(* IEC 61131-3 sources: 89152_FlorisHendrix_AfstudeerProject/89152_FlorisHendrix_ExamenProject/Stations/Terminal/HMI/Network/NewAgeSettings, 1 file *)

(* ---- ONE_NewAgeSettings_Table.st ---- *)
#define OBJECTS_CONFIG

//Define part of class USB_DataExchange
#define USB_DATA_CMD                  16#10
#define USB_DataExchangeBase_Timeout  10ms
#define continue goto LABEL_continue
#include "..\..\Source\interfaces\lsl_st_Usb.h"
//Define part of class DisplaySettings
#define DISPLAYSETTINGS_OS_STARTVERSION_SALAMANDER 0x9100  // salamder starts with v 9.1.00

#define DISPLAYSETTINGS_GRAPHIX_MAX_BRIGHTNESS  255 //(2^8-1) = 255
#define DISPLAYSETTINGS_USB_MAX_BRIGHTNESS      255 //(2^8-1) = 255
#define DISPLAYSETTINGS_MIN_BRIGHTNESS_INPUT      0
#define DISPLAYSETTINGS_MAX_BRIGHTNESS_INPUT    100

#define DISPLAYSETTINGS_MIN_PWM_INPUT          0
#define DISPLAYSETTINGS_MAX_PWM_INPUT          100
#define DISPLAYSETTINGS_PWM_PERIODE_TIME       10000

#define DISPLAYSETTINGS_USB_REQ_TIMER_UP 1000

#define DISPLAYSETTINGS_USB_INIT_ERROR    -1

#define DISPLAYSETTINGS_BRIGHTNESS_ERROR    -1

#define DISPLAYSETTINGS_TASKOBJECT_NOT_FOUND    -5

#define DISPLAYSETTINGS_STATE_OK                0

#define DISPLAYSETTINGS_BACKGROUNDTASK_ERROR    -1
#define DISPLAYSETTINGS_CAN_OBJECT_ERROR        -2
#define DISPLAYSETTINGS_GRAPHIX_ERROR           -3
#define DISPLAYSETTINGS_PSOC_ERROR               -4

#define DISPLAYSETTINGS_BACKLIGHT_SWITCHOFF_TIME 1000 //1 second
#include "..\..\Source\interfaces\lsl_st_kernel.h"
#include "..\..\Source\interfaces\lsl_st_pci.h"
#include "..\..\Source\interfaces\lsl_st_pwm.h"
#include "..\..\Source\interfaces\lsl_st_gpio.h"
#include "..\..\Source\interfaces\lsl_st_screensaver.h"
//Define part of class KeyPadANumStdTemplate
#define KEY_LAYOUT_LINE_1   2#11111111110
#define KEY_LAYOUT_LINE_2   2#11111111110
#define KEY_LAYOUT_LINE_3   2#01111111110
#define KEY_LAYOUT_LINE_4   2#00000000111

#define KEYPAD_ANUM_BUTTON_WIDTH      60
#define KEYPAD_ANUM_BUTTON_HEIGHT     60

#define KEYPAD_ANUM_BUTTON_XOFF       5
#define KEYPAD_ANUM_BUTTON_YOFF       85

#define KEYPAD_ANUM_WIDTH             680
#define KEYPAD_ANUM_HEIGHT            350

#define KEYPAD_ANUM_INPUT_XOFF        5
#define KEYPAD_ANUM_INPUT_YOFF        45
#define KEYPAD_ANUM_INPUT_HEIGHT      30

#define KEYPAD_ANUM_TITLE_XOFF        5
#define KEYPAD_ANUM_TITLE_YOFF        5
#define KEYPAD_ANUM_TITLE_HEIGHT      30

#define KEYPAD_ANUM_ESC_WIDTH         30
//Define part of class KeyPadNumStdTemplate
#define KEYPAD_NUM_BUTTON_WIDTH       80
#define KEYPAD_NUM_BUTTON_HEIGHT      80

#define KEYPAD_NUM_BUTTON_XOFF        5
#define KEYPAD_NUM_BUTTON_YOFF        105

#define KEYPAD_NUM_WIDTH              330
#define KEYPAD_NUM_HEIGHT             435

#define KEYPAD_NUM_INPUT_XOFF         5
#define KEYPAD_NUM_INPUT_YOFF         45
#define KEYPAD_NUM_INPUT_HEIGHT       30

#define KEYPAD_NUM_TITLE_XOFF         7
#define KEYPAD_NUM_TITLE_YOFF         5
#define KEYPAD_NUM_TITLE_HEIGHT       30

#define KEYPAD_NUM_LIMIT_XOFF         5
#define KEYPAD_NUM_LIMIT_YOFF         80
#define KEYPAD_NUM_LIMIT_WIDTH        80
#define KEYPAD_NUM_LIMIT_HEIGTH       20

#define KEYPAD_NUM_UNIT_WIDTH         70
#define KEYPAD_NUM_UNIT_HEIGTH        20

#define KEYPAD_NUM_ESC_WIDTH          30
//Define part of class SystemLogging
//texts for indicating type of loginformation
#define LOG_TYPE_ERROR    ("ERROR:")
#define LOG_TYPE_WARNING  ("WARNING:")
#define LOG_TYPE_DEBUG    ("DEBUG:")
#define LOG_TYPE_INFO     ("INFO:")
//Define part of class TouchCalib
// Default-Settings for the Touch-Calibration
//-------------------------------------------------------------------------------------------------

#define   TouchCalib_UDCVersion                                         1
#define   TouchCalib_NoAnything                                         2

#define   TouchCalib_TextTouchScreen                                    "Please touch the screen to start!"
#define   TouchCalib_TextTouchCrosshair                                 "Please touch the crosshair!"
#define   TouchCalib_TextCalibSuccessful                                "Calibration successful! Please touch the screen to continue."
#define   TouchCalib_TextCalibFailed                                    "Calibration failed! Please touch the screen to calibrate again."
#define   TouchCalib_TextNextScreen                                     "Calibration successful! Please touch the NEXT device to continue."

#define   TouchCalib_TextIdxTouchScreen                                 0
#define   TouchCalib_TextIdxTouchCrosshair                              1
#define   TouchCalib_TextIdxCalibSuccessful                             2
#define   TouchCalib_TextIdxCalibFailed                                 3
#define   TouchCalib_TextIdxNextScreen                                  4

#define   TouchCalib_StdTextAttrib                                      T_SOLID OR T_COPY OR T_PROP

#define   TouchCalib_CrosshairSize                                      40                                            // The length and width of the crosshair (if no image is chosen) [pixel]

#define   TouchCalib_MinTimeBewtweenTouchEvent                         100 ms

FUNCTION GLOBAL TAB ONE_NewAgeSettings
-1$UINT, 0$UINT,
1$UINT, 0$UINT,

15$UDINT,
TO_UDINT(3788417926), "_Global", 0$UINT, 15$UINT, 0$UINT,
TO_UDINT(1108585033), "_LanguageSelection", 0$UINT, 5$UINT, 1$UINT,
TO_UDINT(2980745877), "_MyIO", 0$UINT, 3$UINT, 0$UINT,
TO_UDINT(3599188277), "_Screen", 0$UINT, 3$UINT, 0$UINT,
TO_UDINT(3043040051), "_ScrollArea", 0$UINT, 15$UINT, 0$UINT,
TO_UDINT(2779823616), "_ScrollArea2", 0$UINT, 8$UINT, 0$UINT,
TO_UDINT(3306153856), "DisplaySettings", 1$UINT, 39$UINT, 1$UINT,
TO_UDINT(1679073929), "KeyPadANumStdTemplate", 3$UINT, 0$UINT, 1$UINT,
TO_UDINT(980817768), "KeyPadImagesStdTemplate", 2$UINT, 0$UINT, 2$UINT,
TO_UDINT(1267823535), "KeyPadNumStdTemplate", 1$UINT, 0$UINT, 1$UINT,
TO_UDINT(1903583397), "Ram", 1$UINT, 3$UINT, 1$UINT,
TO_UDINT(3719262472), "ScreenSaver", 1$UINT, 13$UINT, 1$UINT,
TO_UDINT(90452573), "SystemLogging", 1$UINT, 5$UINT, 1$UINT,
TO_UDINT(627189056), "TouchCalib", 1$UINT, 4$UINT, 1$UINT,
TO_UDINT(1659734526), "USB_DataExchange", 1$UINT, 14$UINT, 0$UINT,

_NO_ATTR, TO_UDINT(2359166249), "_LANGUAGESELECTION1",

1$UINT, TO_UDINT(474634808), "SCREENSAVER1\DISPLAYSETTINGS",

_NO_ATTR, TO_UDINT(1679073929), "KEYPADANUMSTDTEMPLATE",

1$UINT, TO_UDINT(860932433), "KEYPADANUMSTDTEMPLATE\KEYPADIMG",
1$UINT, TO_UDINT(1346448759), "KEYPADNUMSTDTEMPLATE\KEYPADIMG",

_NO_ATTR, TO_UDINT(1267823535), "KEYPADNUMSTDTEMPLATE",

_NO_ATTR, TO_UDINT(2623333383), "CLEANSCREENTIME",

_NO_ATTR, TO_UDINT(2379925748), "SCREENSAVER1",

_NO_ATTR, TO_UDINT(2516821708), "SYSTEMLOGGING1",

_NO_ATTR, TO_UDINT(4112894978), "TOUCHCALIB1",

//Internal connections
0$UDINT,
3$UDINT,
TO_UDINT(2), "KeyPadImg", TO_UDINT(3),
TO_UDINT(5), "KeyPadImg", TO_UDINT(4),
TO_UDINT(7), "DisplaySettings", TO_UDINT(1),
0$UDINT,
0$UDINT,

//Initialization values
0$UDINT,
18$UDINT,
TO_UDINT(0), "LineWidth", TO_UDINT(70),//|NewAgeSettings._LanguageSelection1.LineWidth;
TO_UDINT(0), "LineHighness", TO_UDINT(30),//|NewAgeSettings._LanguageSelection1.LineHighness;
TO_UDINT(0), "ExtendedScrollBar", TO_UDINT(0),//|NewAgeSettings._LanguageSelection1.ExtendedScrollBar;
TO_UDINT(0), "Config", TO_UDINT(3),//|NewAgeSettings._LanguageSelection1.Config;
TO_UDINT(1), "Brightness", TO_UDINT(100),//|NewAgeSettings.ScreenSaver1\DisplaySettings.Brightness;
TO_UDINT(1), "ScreensaverTime", TO_UDINT(60),//|NewAgeSettings.ScreenSaver1\DisplaySettings.ScreensaverTime;
TO_UDINT(2), "No", TO_UDINT(_WIN_EDITOR_ANUMERIC),//|NewAgeSettings.KeyPadANumStdTemplate.No;
TO_UDINT(2), "ImA", TO_UDINT(ImA_Window),//|NewAgeSettings.KeyPadANumStdTemplate.ImA;
TO_UDINT(5), "No", TO_UDINT(_WIN_EDITOR_NUMERIC),//|NewAgeSettings.KeyPadNumStdTemplate.No;
TO_UDINT(5), "ImA", TO_UDINT(IMA_WINDOW),//|NewAgeSettings.KeyPadNumStdTemplate.ImA;
TO_UDINT(6), "", TO_UDINT(5),//|NewAgeSettings.CleanScreenTime.Data;
TO_UDINT(7), "sDelayScreenSaver", TO_UDINT(0),//|NewAgeSettings.ScreenSaver1.sDelayScreenSaver;
TO_UDINT(7), "sDelayBacklight", TO_UDINT(0),//|NewAgeSettings.ScreenSaver1.sDelayBacklight;
TO_UDINT(7), "BrightnessMinStart", TO_UDINT(20),//|NewAgeSettings.ScreenSaver1.BrightnessMinStart;
TO_UDINT(8), "ExtLoggingActive", TO_UDINT(TRUE),//|NewAgeSettings.SystemLogging1.ExtLoggingActive;
TO_UDINT(8), "ActivateTrace", TO_UDINT(0),//|NewAgeSettings.SystemLogging1.ActivateTrace;
TO_UDINT(9), "SelectOrderNo", TO_UDINT(-1),//|NewAgeSettings.TouchCalib1.SelectOrderNo;
TO_UDINT(9), "Tolerance", TO_UDINT(20),//|NewAgeSettings.TouchCalib1.Tolerance;

//Symbolic initialization values
0$UDINT,
0$UDINT,

//Initialization of string values
0$UDINT,
0$UDINT,

//Configuration of tasks (RealTime, Cyclic, Background)
0$UDINT,
0$UDINT,

0$UDINT,
0$UDINT,

0$UDINT,
1$UDINT,
TO_UDINT(1), (-1)$UDINT, 4194303$DINT, 	//SCREENSAVER1\DISPLAYSETTINGS

//External connections
0$UDINT,
5$UDINT,
TO_UDINT(0), "Lse", C_DIR, TO_UDINT(299963966), "Lse","Lse",
TO_UDINT(2), "Lse", C_DIR, TO_UDINT(299963966), "Lse","Lse",
TO_UDINT(5), "Lse", C_DIR, TO_UDINT(299963966), "Lse","Lse",
TO_UDINT(7), "Lse", C_DIR, TO_UDINT(299963966), "Lse","Lse",
TO_UDINT(9), "Lse", C_DIR, TO_UDINT(299963966), "Lse","Lse",

//Magic internal connections
0$UDINT,
0$UDINT,

//Configuration of timeslots of tasks (RealTime, Cyclic)
#ifdef __LSLLDR_TIMESLOTS__
0$UDINT,
0$UDINT,

0$UDINT,
0$UDINT,

#endif //__LSLLDR_TIMESLOTS__

//MultiMaster connections
#ifdef __LSLLDR_MULTIMASTER__
0$UDINT,
0$UDINT,
#endif //__LSLLDR_MULTIMASTER__

//Configuration for task ID (RealTime, CyclicTime)
#ifdef __LSLLDR_TASKID__
"\\\\TASKS2  "
0$UDINT,
0$UDINT,

0$UDINT,
0$UDINT,

0$UDINT,
1$UDINT,
(0)$UDINT, 	//SCREENSAVER1\DISPLAYSETTINGS

#endif //__LSLLDR_TASKID__

END_FUNCTION
